// TIA Portal V21 export
// export: Created 2026-08-21T20:18:50.5323427Z, ExportSetting None, DisplayName Totally Integrated Automation Portal, DisplayVersion V21, DisplayName STEP 7 Professional, DisplayVersion V21, DisplayName STEP 7 Safety, DisplayVersion V21, DisplayName Tech WebApplication, DisplayVersion V21, DisplayName WinCC Basic/Comfort/Advanced, DisplayVersion V21, DisplayName WinCC Professional, DisplayVersion V21, DisplayName WinCC Unified, DisplayVersion V21
DATA_BLOCK "Global_Limits_Interlocks"   // DB58
{ S7_Optimized_Access := 'TRUE' }
// stored: MemoryReserve 100
   VAR
      ExternalLevel_Interlock : Real := 2900.0;
      InternalLevel_Interlock : Real := 2700.0;
   END_VAR
BEGIN
END_DATA_BLOCK
